Fanuc KAREL source: kt00146.KL

-- PROVISIONAL review KL for V1013-1; original PC SHA256 6fa442be96b80a219a4a968ecce0f07c6446490535ccae91827d70da4270baa2
-- Incomplete behavior may be omitted. Consult companion uncertainty JSON. Do not deploy.
PROGRAM KT00146
%NOLOCKGROUP
VAR
  I2 : INTEGER
  OUT : REAL
-- UNRESOLVED_DECL Y1 type=002018
BEGIN
  -- UNRESOLVED_PC offsets 5-19; opcodes 2E,22,9D,33,B2
  -- UNRESOLVED_PC offsets 24-35; opcodes 2E,23
  -- UNRESOLVED_PC offsets 40-63; opcodes 22,9D,33,B1,21,55,64,23
  -- UNRESOLVED_PC offsets 68-72; opcodes 7F
END KT00146
